// TIA Portal V20 export
TYPE "Teile Status"
   STRUCT
      "Teil eingelegt" : Bool := 0;
      "Teil IO" : Bool := 0;
      "Teil NIO" : Bool := 0;
      Leer : Bool := 1;
      Reset_Status : Bool := 0;
      "NIO Rundlauf" : Bool;
      "NIO Höhenmessung Pos10" : Bool;
      "NIO Pos9_2" : Bool;
      "NIO Fügen Pos 9_3" : Bool;
      "NIO Bördeln Pos 9_4" : Bool;
      "NIO Messung Pos 9_5" : Bool;
      "NIO Sicken Pos 8_0" : Bool;
      Statuswort : DInt := 0;
   END_STRUCT;
END_TYPE
